(* IEC 61131-3 sources: plcassist-cli/packages/volt-lsp-iec/test-corpus/pro2193/Device/Plc Logic/Application/09 Misc/Library Manager/CAA ResMan, 20 files *)

(* ---- VERSIONCONSTANTS.gvl ---- *)
VAR_GLOBAL
	GC_BYVERSION : BYTE := 1;
	GC_BYVERSION_1 : BYTE := 0;
END_VAR

(* ---- _BLOCKGETDATA.fun ---- *)
FUNCTION _BLOCKGETDATA : CAA.PVOID
VAR_INPUT
	HBLOCK : CAA.HANDLE;
	PEERROR : POINTER TO ERROR;
END_VAR
END_FUNCTION

(* ---- _POOLCREATEP.fun ---- *)
FUNCTION _POOLCREATEP : CAA.HANDLE
VAR_INPUT
	SZBLOCKSIZE : CAA.SIZE;
	SZMEMSIZE : CAA.SIZE;
	PMEMORY : CAA.PVOID;
	EEMPTY : INT;
	PEERROR : POINTER TO ERROR;
END_VAR
END_FUNCTION

(* ---- _POOLDELETE.fun ---- *)
FUNCTION _POOLDELETE : ERROR
VAR_INPUT
	HPOOL : CAA.HANDLE;
END_VAR
END_FUNCTION

(* ---- _POOLEXTENDH.fun ---- *)
FUNCTION _POOLEXTENDH : ERROR
VAR_INPUT
	HPOOL : CAA.HANDLE;
	CTNUMBLOCKS : CAA.COUNT;
END_VAR
END_FUNCTION

(* ---- _POOLGETBLOCK.fun ---- *)
FUNCTION _POOLGETBLOCK : CAA.HANDLE
VAR_INPUT
	HPOOL : CAA.HANDLE;
	PEERROR : POINTER TO ERROR;
END_VAR
END_FUNCTION

(* ---- _POOLPUTBLOCK.fun ---- *)
FUNCTION _POOLPUTBLOCK : ERROR
VAR_INPUT
	HBLOCK : CAA.HANDLE;
END_VAR
END_FUNCTION

(* ---- CHECK.fun ---- *)
FUNCTION CHECK : CAA.HANDLE
VAR_INPUT
	HCHECK : CAA.HANDLE;
	PEERROR : POINTER TO ERROR;
END_VAR
END_FUNCTION

(* ---- CLASSCREATE.fun ---- *)
FUNCTION CLASSCREATE : CAA.HANDLE
VAR_INPUT
	PFUNCTION : CAA.PVOID;
	CTMAXHANDLES : CAA.COUNT;
	PEERROR : POINTER TO ERROR;
END_VAR
END_FUNCTION

(* ---- CLASSDELETE.fun ---- *)
FUNCTION CLASSDELETE : ERROR
VAR_INPUT
	HCLASS : CAA.HANDLE;
END_VAR
END_FUNCTION

(* ---- CLASSFREE.fun ---- *)
FUNCTION CLASSFREE : ERROR
VAR_INPUT
	HCLASS : CAA.HANDLE;
END_VAR
END_FUNCTION

(* ---- GETCLASS.fun ---- *)
FUNCTION GETCLASS : CAA.HANDLE
VAR_INPUT
	HCHECK : CAA.HANDLE;
	PEERROR : POINTER TO ERROR;
END_VAR
END_FUNCTION

(* ---- GETCLASSINFO.fun ---- *)
FUNCTION GETCLASSINFO : ERROR
VAR_INPUT
	HCLASS : CAA.HANDLE;
	PCLASSINFO : POINTER TO CLASS_INFO;
END_VAR
END_FUNCTION

(* ---- GETINFO.fun ---- *)
FUNCTION GETINFO : ERROR
VAR_INPUT
	PINFO : POINTER TO INFO;
END_VAR
END_FUNCTION

(* ---- GETPARENT.fun ---- *)
FUNCTION GETPARENT : CAA.HANDLE
VAR_INPUT
	HCHECK : CAA.HANDLE;
	PEERROR : POINTER TO ERROR;
END_VAR
END_FUNCTION

(* ---- GETSUPPLIERVERSION.fun ---- *)
FUNCTION GETSUPPLIERVERSION : WORD
VAR_INPUT
	XDUMMY : BOOL;
END_VAR
END_FUNCTION

(* ---- REGISTER.fun ---- *)
FUNCTION REGISTER : CAA.HANDLE
VAR_INPUT
	HCLASS : CAA.HANDLE;
	HRESSOURCE : CAA.HANDLE;
	PEERROR : POINTER TO ERROR;
END_VAR
END_FUNCTION

(* ---- SETPARENT.fun ---- *)
FUNCTION SETPARENT : ERROR
VAR_INPUT
	HCHECK : CAA.HANDLE;
	HCHECKPARENT : CAA.HANDLE;
END_VAR
END_FUNCTION

(* ---- UNREGISTER.fun ---- *)
FUNCTION UNREGISTER : ERROR
VAR_INPUT
	HCHECK : CAA.HANDLE;
END_VAR
END_FUNCTION

(* ---- RSMCLASS.fb ---- *)
FUNCTION_BLOCK RSMCLASS
VAR
	_HPOOL : CAA.HANDLE;
	_ADWPOOL : ARRAY [0..19] OF __XWORD;
	_PLIST : POINTER TO RSM_HANDLE;
END_VAR
END_FUNCTION_BLOCK

METHOD FB_EXIT : BOOL
VAR_INPUT
	BINCOPYCODE : BOOL;
END_VAR
END_METHOD

METHOD REGISTER : CAA.HANDLE
VAR_INPUT
	HHANDLE : CAA.HANDLE;
	PEERROR : POINTER TO ERROR;
END_VAR
END_METHOD

METHOD CLOSE : ERROR
VAR_INPUT
	HHANDLE : CAA.HANDLE;
END_VAR
END_METHOD

METHOD SEARCH : CAA.HANDLE
VAR_INPUT
	HHANDLE : CAA.HANDLE;
END_VAR
END_METHOD

METHOD UNREGISTER : ERROR
VAR_INPUT
	HHANDLE : CAA.HANDLE;
END_VAR
END_METHOD

METHOD FB_INIT : BOOL
VAR_INPUT
	BINITRETAINS : BOOL;
	BINCOPYCODE : BOOL;
END_VAR
END_METHOD

METHOD TRANSLATE : CAA.HANDLE
VAR_INPUT
	HHANDLE : CAA.HANDLE;
END_VAR
VAR_OUTPUT
	EERROR : ERROR;
END_VAR
END_METHOD
